(* IEC 61131-3 sources: ISA-88-Bioreactor-Automation-Template-DE-IE/ISA-88-Bioreactor-Automation-Template-DE-IE.fbsdev/CycleManager.iecapp^, 2 files *)

(* ---- CycleManager_FB_ST.fb.st ---- *)
FUNCTION_BLOCK CycleManager_FB_ST
VAR_INPUT
    Global_Start        : BOOL;   // Operator command to start plant
    Global_Stop         : BOOL;   // Operator command to stop plant
    Tank1_CycleComplete : BOOL;   // Tank 1 cycle finished
    Tank2_CycleComplete : BOOL;   // Tank 2 cycle finished
    CIP_Complete_T1     : BOOL;   // Tank 1 CIP finished
    CIP_Complete_T2     : BOOL;   // Tank 2 CIP finished
    Utilities_OK        : BOOL;   // Consolidated utility status
    Interlock_OK        : BOOL;   // Consolidated interlock status
END_VAR

VAR_OUTPUT
    Plant_Active     : BOOL := FALSE; // Plant running
    Plant_Stopped    : BOOL := TRUE;  // Plant stopped
    Tank1_StartCycle : BOOL := FALSE; // Command to start Tank 1 cycle
    Tank2_StartCycle : BOOL := FALSE; // Command to start Tank 2 cycle
    Tank1_StartCIP   : BOOL := FALSE; // Command to start Tank 1 CIP
    Tank2_StartCIP   : BOOL := FALSE; // Command to start Tank 2 CIP
END_VAR

VAR
    Tank1_NeedsCIP : BOOL := FALSE;
    Tank2_NeedsCIP : BOOL := FALSE;
END_VAR

// Plant start/stop logic
IF Global_Start AND Utilities_OK AND Interlock_OK THEN
    Plant_Active := TRUE;
    Plant_Stopped := FALSE;
END_IF;

IF Global_Stop THEN
    Plant_Active := FALSE;
    Plant_Stopped := TRUE;
    Tank1_StartCycle := FALSE;
    Tank2_StartCycle := FALSE;
    Tank1_StartCIP := FALSE;
    Tank2_StartCIP := FALSE;
END_IF;

// Tank 1 cycle/CIP orchestration
IF Plant_Active THEN
    IF Tank1_CycleComplete THEN
        Tank1_NeedsCIP := TRUE;
    END_IF;

    IF Tank1_NeedsCIP AND NOT Tank1_StartCycle THEN
        Tank1_StartCIP := TRUE;
    END_IF;

    IF CIP_Complete_T1 THEN
        Tank1_NeedsCIP := FALSE;
        Tank1_StartCIP := FALSE;
        Tank1_StartCycle := TRUE; // Ready for next production cycle
    END_IF;
END_IF;

// Tank 2 cycle/CIP orchestration
IF Plant_Active THEN
    IF Tank2_CycleComplete THEN
        Tank2_NeedsCIP := TRUE;
    END_IF;

    IF Tank2_NeedsCIP AND NOT Tank2_StartCycle THEN
        Tank2_StartCIP := TRUE;
    END_IF;

    IF CIP_Complete_T2 THEN
        Tank2_NeedsCIP := FALSE;
        Tank2_StartCIP := FALSE;
        Tank2_StartCycle := TRUE; // Ready for next production cycle
    END_IF;
END_IF;

(* ---- PLC_PRG.prg.st ---- *)
PROGRAM PLC_PRG
VAR
    // Supervisory
    CycleMgr      : CycleManager_FB_ST;

    // Submodules
    TankCycle     : TankCycler_FB_ST;
    PumpCtrl      : PumpController_FB_ST;
    ThermalCtrl   : ThermalManager_FB_ST;
    MixerCtrl     : MixerController_FB_ST;
    CIPCtrl       : CIPManager_FB_ST;
    AlarmCtrl     : AlarmCtrl_FB_ST;
    InterlockCtrl : InterlockManager_FB_ST;
    UtilityCtrl   : UtilityMonitor_FB_ST;
    BatchCtrl     : BatchCounter_FB_ST;

    // Operator inputs
    Global_Start  : BOOL;
    Global_Stop   : BOOL;

    // Supervisory outputs
    Plant_Active     : BOOL;
    Plant_Stopped    : BOOL;
    Tank1_StartCycle : BOOL;
    Tank1_StartCIP   : BOOL;
END_VAR

// --- Supervisory orchestration ---
CycleMgr(
    Global_Start := Global_Start,
    Global_Stop := Global_Stop,
    Tank1_CycleComplete := TankCycle.Cycle_Complete,
    Tank2_CycleComplete := FALSE, // add if you have Tank2
    CIP_Complete_T1 := CIPCtrl.CIP_Complete,
    CIP_Complete_T2 := FALSE,
    Utilities_OK := UtilityCtrl.Utilities_OK,
    Interlock_OK := InterlockCtrl.Interlock_OK,
    Plant_Active => Plant_Active,
    Plant_Stopped => Plant_Stopped,
    Tank1_StartCycle => Tank1_StartCycle,
    Tank1_StartCIP => Tank1_StartCIP
);

// --- Submodules execution ---
TankCycle(
    Start_Cycle := Tank1_StartCycle,
    Stop_Cycle := Global_Stop,
    T1_Level_High := T1_Level_High,
    T1_Level_Low := T1_Level_Low,
    T1_Temp_Sensor := T1_Temp_Sensor,
    T1_Temp_Setpoint := T1_Temp_Setpoint
);

PumpCtrl(
    Cycle_Active := TankCycle.Cycle_Active,
    Discharge_Complete := TankCycle.Discharge_Complete
);

ThermalCtrl(
    Cycle_Active := TankCycle.Cycle_Active,
    Mix_Complete := TankCycle.Mix_Complete,
    Tn_Temp_Value := T1_Temp_Sensor,
    Tn_Temp_Setpoint := T1_Temp_Setpoint
);

MixerCtrl(
    Cycle_Active := TankCycle.Cycle_Active,
    Fill_Complete := TankCycle.Fill_Complete
);

CIPCtrl(
    Start_CIP := Tank1_StartCIP,
    Cycle_Complete := TankCycle.Cycle_Complete
);

AlarmCtrl(
    Pump_Alarm := PumpCtrl.Pump_Alarm,
    Thermal_Alarm := ThermalCtrl.Thermal_Alarm,
    Mixer_Alarm := MixerCtrl.Mixer_Alarm,
    CIP_Alarm := CIPCtrl.CIP_Alarm,
    Ack_Alarm := Ack_Alarm
);

InterlockCtrl(
    Cycle_Active := TankCycle.Cycle_Active,
    Utility_OK := UtilityCtrl.Utilities_OK
);

UtilityCtrl(); // monitors steam, water, air

BatchCtrl(
    Cycle_Complete := TankCycle.Cycle_Complete,
    Reset_Counter := Reset_Counter
);
